{attribute 'pack_mode' := '1'}
TYPE ST_AirConditionerPublishData :
STRUCT
	Header		:	ST_MqttHeader;
	Devices		:	ARRAY[0..GVL_PARAM.AIR_CONDITIONER_COUNT-1] OF ST_AirConditionerPublish_V1;
END_STRUCT
END_TYPE

(* stored: Version 1.1.0.1, ProductVersion 3.1.4024.15
   DUT ST_AirConditionerPublishData: Id {97fe4731-03ca-4fa7-8100-ebd10c3ac884} *)
